Fanuc KAREL source: KA00086.KL

PROGRAM KA00086
%NOLOCKGROUP
VAR
  SRC: JOINTPOS
  DST: REAL
BEGIN
  DST = SRC
END KA00086
